Fanuc KAREL source: kd00047.KL

PROGRAM KD00047
%STACKSIZE=65535
%PRIORITY=65535
%NOLOCKGROUP
VAR
I : INTEGER
J : INTEGER
B : BOOLEAN
R : REAL
S : STRING[80]
V : VECTOR
BEGIN
V.X=1.0
-- UNRESOLVED_PC line 13 opcodes [01 49 2E 0A 82 0B] marker_code=20
END KD00047
